Universal Robots PolyScope program: example.urp

Program tanghua_template (installation=default directory=/programs/usbdisk createdIn=3.15.6.0 lastSavedIn=3.15.8.106339)
Calibrated DH parameters: a=[0, -0.425, -0.3922, 0, 0, 0]; d=[0.1625, 0, 0, 0.1333, 0.0997, 0.0996]; alpha=[1.570796, 0, 0, 1.570796, -1.570796, 0]; deltaTheta=[0, 0, 0, 0, 0, 0]
Robot Program (runOnlyOnce=true)
  Script file example.script
    | def Program():
    | end
    | Program()
